// TIA Portal V21 export
// export: Created 2026-11-10T19:16:48.7645305Z, ExportSetting WithDefaults, DisplayName Totally Integrated Automation Portal, DisplayVersion V21 Update 3, DisplayName STEP 7 Professional, DisplayVersion V21 Update 3, DisplayName STEP 7 Safety, DisplayVersion V21, DisplayName Tech WebApplication, DisplayVersion V21, DisplayName WinCC Basic/Comfort/Advanced, DisplayVersion V21 Update 3, DisplayName WinCC Unified, DisplayVersion V21 Update 3
DATA_BLOCK "DB_NonOpt"   // DB7
{ S7_Optimized_Access := 'FALSE' }
VERSION : 0.1
// stored: AutoNumber true, DBAccessibleFromOPCUA true, DBAccessibleFromWebserver true, IsOnlyStoredInLoadMemory false, IsWriteProtectedInAS false
   VAR RETAIN
      b0 : Bool;
      b1 : Bool;
      "by" : Byte;
      i : Int := 5;
      d : DInt;
      r : Real;
      t : Time;
      "dt" : Date_And_Time;
      s : String[12] := 'std';
      arr : Array[1..4] of Word;
      "m" : Array[0..1, 0..2] of Int;
      st : Struct
         x : Bool;
         y { ExternalWritable := 'False'} : Real := 2.5;
      END_STRUCT;
      u { S7_SetPoint := 'True'} : "UDT_Inner";
   END_VAR
BEGIN
   "m"[1,2] := -3;
END_DATA_BLOCK
